(* IEC 61131-3 sources: 2026_Projet_YGO_ExcavatriceDragage/TOOLS/TEST_AUTO_CI/RESULTS/C_DIAG_RESEAUX/tests, 4 files *)

(* ---- test_fb_autoresettransientdiag.st ---- *)
(* =========================================================================
   FB_AutoResetTransientDiag — preuve isolee (T352, parent T278)
   =========================================================================
   Pourquoi ce fichier existe : T278 a livre le FB et son cablage SANS aucun
   test unitaire, et ses deux entrees d'autorisation StartupEnable /
   PowerRearmEnable ont ete cablees sur deux booleens d'une GVL de simulation
   valant FALSE par defaut et sans aucun ecrivain (PRG_02_Acquisition.st:225-226,
   GVL_Simulation.st:106-107). Consequence mesuree sur machine reelle : State
   reste bloque a 0, Phase ne passe jamais a 1 ni a 2, ResetPulse ne bouge
   jamais. Ces cas prouvent que la logique INTERNE du FB est saine des que les
   deux entrees valent TRUE — le defaut etait donc bien en amont du FB.

   Identifiants TC-T352-xxx : cas d'execution rattaches a la tache T352. Ils ne
   prennent AUCUN identifiant TC-P12 du catalogue AF-12 : ce catalogue s'arrete
   a TC-P12-050 et un TC-P12-060 a ete explicitement REFUSE par l'humain
   (AF_Partie-12_Fonction_Diagnostic_v1.4.md, ligne 348).

   Ce fichier prouve des comportements OBSERVABLES par les sorties publiques
   (ResetPulse, SequenceActive, Lockout, Cancelled, Phase, AttemptCount) :
   State et StartupStarted sont des VAR privees, non lisibles de l'exterieur.

   Gardes de securite couvertes, jamais affaiblies :
     FB_AutoResetTransientDiag.st:70  SafeCommon = EmergencyChainClosed AND
                                      NOT PowerCutOffActive AND NOT MotionActive
     FB_AutoResetTransientDiag.st:122 annulation immediate si SafeCommon tombe
   ========================================================================= *)

SETUP
VAR
    FB : FB_AutoResetTransientDiag;
END_VAR
END_SETUP

(* -------------------------------------------------------------------------
   Cas nominal : demarrage, stabilisation, impulsion unique, verrouillage.
   C'est exactement le scenario que l'observateur ne voyait jamais sur machine.
   ------------------------------------------------------------------------- *)
TEST 'TC-T352-001 Demarrage par defaut : Phase 1, impulsion apres stabilisation, verrouillage'
    (* Scan 0 : conditions nominales, contacteur au repos -> la sequence demarre *)
    FB(Enable := TRUE,
       StartupEnable := TRUE,
       PowerRearmEnable := TRUE,
       EmergencyChainClosed := TRUE,
       PowerContactorEngaged := FALSE,
       PowerCutOffActive := FALSE,
       MotionActive := FALSE,
       DiagnosticsStable := TRUE,
       Cfg_MaxAttempts := 1,
       Cfg_StabilizationTime := T#1s,
       Cfg_InterAttemptTime := T#1s);
    ASSERT_TRUE(FB.SequenceActive, 'StartupEnable=TRUE -> sequence active des le 1er scan');
    ASSERT_EQ(FB.Phase, 1, 'Phase 1 = sequence de demarrage engagee');

    (* Scan 1 : aucune impulsion, la stabilisation est en cours *)
    FB(Enable := TRUE, StartupEnable := TRUE, PowerRearmEnable := TRUE,
       EmergencyChainClosed := TRUE, PowerContactorEngaged := FALSE,
       PowerCutOffActive := FALSE, MotionActive := FALSE, DiagnosticsStable := TRUE,
       Cfg_MaxAttempts := 1, Cfg_StabilizationTime := T#1s, Cfg_InterAttemptTime := T#1s);
    ASSERT_FALSE(FB.ResetPulse, 'Aucune impulsion avant Cfg_StabilizationTime');

    (* Scan 2 : 1 s ecoulee -> impulsion unique puis verrouillage (MaxAttempts=1) *)
    ADVANCE_TIME(1000000000);
    FB(Enable := TRUE, StartupEnable := TRUE, PowerRearmEnable := TRUE,
       EmergencyChainClosed := TRUE, PowerContactorEngaged := FALSE,
       PowerCutOffActive := FALSE, MotionActive := FALSE, DiagnosticsStable := TRUE,
       Cfg_MaxAttempts := 1, Cfg_StabilizationTime := T#1s, Cfg_InterAttemptTime := T#1s);
    ASSERT_TRUE(FB.ResetPulse, 'Apres 1 s de stabilisation -> ResetPulse=TRUE');
    ASSERT_EQ(FB.AttemptCount, 1, 'Une seule impulsion emise');
    ASSERT_TRUE(FB.Lockout, 'MaxAttempts=1 atteint -> Lockout=TRUE');
    ASSERT_EQ(FB.Phase, 3, 'Phase 3 = salve terminee, attente d''un nouvel evenement');

    (* Scan 3 : impulsion d'un seul scan, puis retour au repos verrouille *)
    FB(Enable := TRUE, StartupEnable := TRUE, PowerRearmEnable := TRUE,
       EmergencyChainClosed := TRUE, PowerContactorEngaged := FALSE,
       PowerCutOffActive := FALSE, MotionActive := FALSE, DiagnosticsStable := TRUE,
       Cfg_MaxAttempts := 1, Cfg_StabilizationTime := T#1s, Cfg_InterAttemptTime := T#1s);
    ASSERT_FALSE(FB.ResetPulse, 'ResetPulse est impulsionnel : FALSE au scan suivant');
    ASSERT_TRUE(FB.Lockout, 'Lockout persiste apres la salve');
    ASSERT_FALSE(FB.SequenceActive, 'Sequence terminee');
END_TEST

(* -------------------------------------------------------------------------
   Le second chemin d'entree, inerte tant que PowerRearmEnable valait FALSE :
   phase 2 declenchee EXCLUSIVEMENT sur front du retour contacteur.
   ------------------------------------------------------------------------- *)
TEST 'TC-T352-002 Post-rearmement : Phase 2 sur front contacteur, impulsion puis verrouillage'
    (* Scan 0 : contacteur au repos, phase demarrage volontairement desactivee *)
    FB(Enable := TRUE,
       StartupEnable := FALSE,
       PowerRearmEnable := TRUE,
       EmergencyChainClosed := TRUE,
       PowerContactorEngaged := FALSE,
       PowerCutOffActive := FALSE,
       MotionActive := FALSE,
       DiagnosticsStable := TRUE,
       Cfg_MaxAttempts := 1,
       Cfg_StabilizationTime := T#1s,
       Cfg_InterAttemptTime := T#1s);
    ASSERT_FALSE(FB.SequenceActive, 'Aucun evenement -> sequence au repos');

    (* Scan 1 : front montant du contacteur -> phase post-rearmement *)
    FB(Enable := TRUE, StartupEnable := FALSE, PowerRearmEnable := TRUE,
       EmergencyChainClosed := TRUE, PowerContactorEngaged := TRUE,
       PowerCutOffActive := FALSE, MotionActive := FALSE, DiagnosticsStable := TRUE,
       Cfg_MaxAttempts := 1, Cfg_StabilizationTime := T#1s, Cfg_InterAttemptTime := T#1s);
    ASSERT_TRUE(FB.SequenceActive, 'Front contacteur -> sequence post-rearmement engagee');
    ASSERT_EQ(FB.Phase, 2, 'Phase 2 = sequence post-rearmement');
    ASSERT_FALSE(FB.ResetPulse, 'Impulsion differee apres stabilisation');

    (* Scan 2 : stabilisation ecoulee -> impulsion puis verrouillage *)
    ADVANCE_TIME(1000000000);
    FB(Enable := TRUE, StartupEnable := FALSE, PowerRearmEnable := TRUE,
       EmergencyChainClosed := TRUE, PowerContactorEngaged := TRUE,
       PowerCutOffActive := FALSE, MotionActive := FALSE, DiagnosticsStable := TRUE,
       Cfg_MaxAttempts := 1, Cfg_StabilizationTime := T#1s, Cfg_InterAttemptTime := T#1s);
    ASSERT_TRUE(FB.ResetPulse, 'Apres stabilisation post-rearmement -> ResetPulse=TRUE');
    ASSERT_EQ(FB.AttemptCount, 1, 'Une impulsion emise');
    ASSERT_TRUE(FB.Lockout, 'Salve epuisee -> Lockout=TRUE');
END_TEST

(* -------------------------------------------------------------------------
   Gardes de securite : aucune impulsion ne doit sortir. Les trois composantes
   de SafeCommon sont testees separement, chacune suffit a interdire la salve.
   ------------------------------------------------------------------------- *)
TEST 'TC-T352-003 Gardes safety : chaine AU ouverte, coupure puissance, mouvement actif'
    (* Chaine AU ouverte : EmergencyChainClosed=FALSE *)
    FB(Enable := TRUE, StartupEnable := TRUE, PowerRearmEnable := TRUE,
       EmergencyChainClosed := FALSE, PowerContactorEngaged := FALSE,
       PowerCutOffActive := FALSE, MotionActive := FALSE, DiagnosticsStable := TRUE,
       Cfg_MaxAttempts := 3, Cfg_StabilizationTime := T#1s, Cfg_InterAttemptTime := T#1s);
    ASSERT_FALSE(FB.SequenceActive, 'Chaine AU ouverte -> aucune sequence');
    ASSERT_FALSE(FB.ResetPulse, 'Chaine AU ouverte -> aucune impulsion');

    (* Coupure puissance active : PowerCutOffActive=TRUE *)
    FB(Enable := TRUE, StartupEnable := TRUE, PowerRearmEnable := TRUE,
       EmergencyChainClosed := TRUE, PowerContactorEngaged := FALSE,
       PowerCutOffActive := TRUE, MotionActive := FALSE, DiagnosticsStable := TRUE,
       Cfg_MaxAttempts := 3, Cfg_StabilizationTime := T#1s, Cfg_InterAttemptTime := T#1s);
    ASSERT_FALSE(FB.SequenceActive, 'Coupure puissance active -> aucune sequence');

    (* Mouvement actif : MotionActive=TRUE *)
    FB(Enable := TRUE, StartupEnable := TRUE, PowerRearmEnable := TRUE,
       EmergencyChainClosed := TRUE, PowerContactorEngaged := FALSE,
       PowerCutOffActive := FALSE, MotionActive := TRUE, DiagnosticsStable := TRUE,
       Cfg_MaxAttempts := 3, Cfg_StabilizationTime := T#1s, Cfg_InterAttemptTime := T#1s);
    ASSERT_FALSE(FB.SequenceActive, 'Mouvement actif -> aucune sequence');

    (* Le temps qui passe ne force rien : meme apres 5 s, toujours aucune impulsion *)
    ADVANCE_TIME(5000000000);
    FB(Enable := TRUE, StartupEnable := TRUE, PowerRearmEnable := TRUE,
       EmergencyChainClosed := TRUE, PowerContactorEngaged := FALSE,
       PowerCutOffActive := FALSE, MotionActive := TRUE, DiagnosticsStable := TRUE,
       Cfg_MaxAttempts := 3, Cfg_StabilizationTime := T#1s, Cfg_InterAttemptTime := T#1s);
    ASSERT_FALSE(FB.ResetPulse, 'Garde safety invalide -> ResetPulse reste FALSE malgre le temps');
    ASSERT_EQ(FB.AttemptCount, 0, 'Aucune tentative consommee sous garde invalide');

    (* Diagnostics reseau instables : la stabilisation ne progresse pas *)
    FB(Enable := TRUE, StartupEnable := TRUE, PowerRearmEnable := TRUE,
       EmergencyChainClosed := TRUE, PowerContactorEngaged := FALSE,
       PowerCutOffActive := FALSE, MotionActive := FALSE, DiagnosticsStable := FALSE,
       Cfg_MaxAttempts := 3, Cfg_StabilizationTime := T#1s, Cfg_InterAttemptTime := T#1s);
    ASSERT_EQ(FB.Phase, 1, 'Sequence engagee mais bloquee en phase 1');
    ADVANCE_TIME(5000000000);
    FB(Enable := TRUE, StartupEnable := TRUE, PowerRearmEnable := TRUE,
       EmergencyChainClosed := TRUE, PowerContactorEngaged := FALSE,
       PowerCutOffActive := FALSE, MotionActive := FALSE, DiagnosticsStable := FALSE,
       Cfg_MaxAttempts := 3, Cfg_StabilizationTime := T#1s, Cfg_InterAttemptTime := T#1s);
    ASSERT_FALSE(FB.ResetPulse, 'Diagnostics instables -> aucune impulsion');
    ASSERT_EQ(FB.AttemptCount, 0, 'Aucune tentative consommee sans diagnostics stables');
END_TEST

(* -------------------------------------------------------------------------
   Annulation en cours de sequence : la garde retombe pendant la salve.
   ------------------------------------------------------------------------- *)
TEST 'TC-T352-004 Annulation : chute de la garde pendant la sequence -> Cancelled + Lockout'
    FB(Enable := TRUE, StartupEnable := TRUE, PowerRearmEnable := TRUE,
       EmergencyChainClosed := TRUE, PowerContactorEngaged := FALSE,
       PowerCutOffActive := FALSE, MotionActive := FALSE, DiagnosticsStable := TRUE,
       Cfg_MaxAttempts := 3, Cfg_StabilizationTime := T#1s, Cfg_InterAttemptTime := T#1s);
    ASSERT_EQ(FB.Phase, 1, 'Sequence engagee');

    (* L'AU s'ouvre pendant la salve -> annulation immediate *)
    ADVANCE_TIME(500000000);
    FB(Enable := TRUE, StartupEnable := TRUE, PowerRearmEnable := TRUE,
       EmergencyChainClosed := FALSE, PowerContactorEngaged := FALSE,
       PowerCutOffActive := FALSE, MotionActive := FALSE, DiagnosticsStable := TRUE,
       Cfg_MaxAttempts := 3, Cfg_StabilizationTime := T#1s, Cfg_InterAttemptTime := T#1s);
    ASSERT_TRUE(FB.Cancelled, 'Garde tombee en cours de sequence -> Cancelled=TRUE');
    ASSERT_TRUE(FB.Lockout, 'Salve annulee -> Lockout=TRUE');
    ASSERT_FALSE(FB.ResetPulse, 'Annulation -> aucune impulsion');
    ASSERT_FALSE(FB.SequenceActive, 'Sequence interrompue');
    ASSERT_EQ(FB.Phase, 3, 'Phase 3 = verrouillage apres annulation');
END_TEST

(* -------------------------------------------------------------------------
   Borne haute : 3 impulsions espacees de Cfg_InterAttemptTime, puis lockout.
   Cadence reelle du FB : impulsion (etat 3) -> scan d'intervalle (retour etat 1)
   -> redemarrage de la stabilisation -> impulsion suivante.
   ------------------------------------------------------------------------- *)
TEST 'TC-T352-005 Borne haute : 3 impulsions espacees puis verrouillage definitif'
    FB(Enable := TRUE, StartupEnable := TRUE, PowerRearmEnable := TRUE,
       EmergencyChainClosed := TRUE, PowerContactorEngaged := FALSE,
       PowerCutOffActive := FALSE, MotionActive := FALSE, DiagnosticsStable := TRUE,
       Cfg_MaxAttempts := 3, Cfg_StabilizationTime := T#1s, Cfg_InterAttemptTime := T#1s);
    ASSERT_EQ(FB.Phase, 1, 'Sequence engagee');

    (* Impulsion 1 *)
    ADVANCE_TIME(1000000000);
    FB(Enable := TRUE, StartupEnable := TRUE, PowerRearmEnable := TRUE,
       EmergencyChainClosed := TRUE, PowerContactorEngaged := FALSE,
       PowerCutOffActive := FALSE, MotionActive := FALSE, DiagnosticsStable := TRUE,
       Cfg_MaxAttempts := 3, Cfg_StabilizationTime := T#1s, Cfg_InterAttemptTime := T#1s);
    ASSERT_TRUE(FB.ResetPulse, 'Impulsion 1 sur 3');
    ASSERT_EQ(FB.AttemptCount, 1, 'Compteur a 1');
    ASSERT_FALSE(FB.Lockout, 'Salve non epuisee -> aucun verrouillage');

    (* Intervalle : la tempo inter-impulsions ramene la sequence en phase 1 *)
    ADVANCE_TIME(1000000000);
    FB(Enable := TRUE, StartupEnable := TRUE, PowerRearmEnable := TRUE,
       EmergencyChainClosed := TRUE, PowerContactorEngaged := FALSE,
       PowerCutOffActive := FALSE, MotionActive := FALSE, DiagnosticsStable := TRUE,
       Cfg_MaxAttempts := 3, Cfg_StabilizationTime := T#1s, Cfg_InterAttemptTime := T#1s);
    ASSERT_FALSE(FB.ResetPulse, 'Intervalle inter-impulsions respecte');
    ASSERT_EQ(FB.AttemptCount, 1, 'Compteur inchange pendant l''intervalle');
    ASSERT_EQ(FB.Phase, 1, 'Retour en phase 1 pour la tentative suivante');

    (* Redemarrage de la stabilisation puis impulsion 2 *)
    ADVANCE_TIME(1000000000);
    FB(Enable := TRUE, StartupEnable := TRUE, PowerRearmEnable := TRUE,
       EmergencyChainClosed := TRUE, PowerContactorEngaged := FALSE,
       PowerCutOffActive := FALSE, MotionActive := FALSE, DiagnosticsStable := TRUE,
       Cfg_MaxAttempts := 3, Cfg_StabilizationTime := T#1s, Cfg_InterAttemptTime := T#1s);
    ASSERT_FALSE(FB.ResetPulse, 'Stabilisation redemarree : pas d''impulsion immediate');

    ADVANCE_TIME(1000000000);
    FB(Enable := TRUE, StartupEnable := TRUE, PowerRearmEnable := TRUE,
       EmergencyChainClosed := TRUE, PowerContactorEngaged := FALSE,
       PowerCutOffActive := FALSE, MotionActive := FALSE, DiagnosticsStable := TRUE,
       Cfg_MaxAttempts := 3, Cfg_StabilizationTime := T#1s, Cfg_InterAttemptTime := T#1s);
    ASSERT_TRUE(FB.ResetPulse, 'Impulsion 2 sur 3');
    ASSERT_EQ(FB.AttemptCount, 2, 'Compteur a 2');
    ASSERT_FALSE(FB.Lockout, 'Salve non epuisee -> aucun verrouillage');

    (* Intervalle puis impulsion 3, qui sature la borne *)
    ADVANCE_TIME(1000000000);
    FB(Enable := TRUE, StartupEnable := TRUE, PowerRearmEnable := TRUE,
       EmergencyChainClosed := TRUE, PowerContactorEngaged := FALSE,
       PowerCutOffActive := FALSE, MotionActive := FALSE, DiagnosticsStable := TRUE,
       Cfg_MaxAttempts := 3, Cfg_StabilizationTime := T#1s, Cfg_InterAttemptTime := T#1s);
    ASSERT_FALSE(FB.ResetPulse, 'Intervalle inter-impulsions respecte (2)');

    ADVANCE_TIME(1000000000);
    FB(Enable := TRUE, StartupEnable := TRUE, PowerRearmEnable := TRUE,
       EmergencyChainClosed := TRUE, PowerContactorEngaged := FALSE,
       PowerCutOffActive := FALSE, MotionActive := FALSE, DiagnosticsStable := TRUE,
       Cfg_MaxAttempts := 3, Cfg_StabilizationTime := T#1s, Cfg_InterAttemptTime := T#1s);
    ASSERT_FALSE(FB.ResetPulse, 'Stabilisation redemarree : pas d''impulsion immediate (2)');

    ADVANCE_TIME(1000000000);
    FB(Enable := TRUE, StartupEnable := TRUE, PowerRearmEnable := TRUE,
       EmergencyChainClosed := TRUE, PowerContactorEngaged := FALSE,
       PowerCutOffActive := FALSE, MotionActive := FALSE, DiagnosticsStable := TRUE,
       Cfg_MaxAttempts := 3, Cfg_StabilizationTime := T#1s, Cfg_InterAttemptTime := T#1s);
    ASSERT_TRUE(FB.ResetPulse, 'Impulsion 3 sur 3');
    ASSERT_EQ(FB.AttemptCount, 3, 'Compteur a 3');
    ASSERT_TRUE(FB.Lockout, 'Borne haute atteinte -> verrouillage');
    ASSERT_EQ(FB.Phase, 3, 'Phase 3 apres salve complete');

    (* Le temps ne relance rien : seul un nouvel evenement rearme la salve *)
    ADVANCE_TIME(10000000000);
    FB(Enable := TRUE, StartupEnable := TRUE, PowerRearmEnable := TRUE,
       EmergencyChainClosed := TRUE, PowerContactorEngaged := FALSE,
       PowerCutOffActive := FALSE, MotionActive := FALSE, DiagnosticsStable := TRUE,
       Cfg_MaxAttempts := 3, Cfg_StabilizationTime := T#1s, Cfg_InterAttemptTime := T#1s);
    ASSERT_FALSE(FB.ResetPulse, 'Aucune 4e impulsion');
    ASSERT_EQ(FB.AttemptCount, 3, 'Compteur fige a la borne');
    ASSERT_TRUE(FB.Lockout, 'Verrouillage conserve');
END_TEST

(* -------------------------------------------------------------------------
   Neutralisation : Enable=FALSE remet le service au repos.
   ------------------------------------------------------------------------- *)
TEST 'TC-T352-006 Neutralisation : Enable=FALSE -> service remis au repos'
    FB(Enable := TRUE, StartupEnable := TRUE, PowerRearmEnable := TRUE,
       EmergencyChainClosed := TRUE, PowerContactorEngaged := FALSE,
       PowerCutOffActive := FALSE, MotionActive := FALSE, DiagnosticsStable := TRUE,
       Cfg_MaxAttempts := 3, Cfg_StabilizationTime := T#1s, Cfg_InterAttemptTime := T#1s);
    ASSERT_TRUE(FB.SequenceActive, 'Sequence engagee avant neutralisation');

    FB(Enable := FALSE, StartupEnable := TRUE, PowerRearmEnable := TRUE,
       EmergencyChainClosed := TRUE, PowerContactorEngaged := FALSE,
       PowerCutOffActive := FALSE, MotionActive := FALSE, DiagnosticsStable := TRUE,
       Cfg_MaxAttempts := 3, Cfg_StabilizationTime := T#1s, Cfg_InterAttemptTime := T#1s);
    ASSERT_FALSE(FB.SequenceActive, 'Enable=FALSE -> sequence neutralisee');
    ASSERT_FALSE(FB.Lockout, 'Enable=FALSE -> verrouillage efface');
    ASSERT_EQ(FB.Phase, 0, 'Enable=FALSE -> retour au repos');
    ASSERT_EQ(FB.AttemptCount, 0, 'Enable=FALSE -> compteur remis a zero');
    ASSERT_FALSE(FB.ResetPulse, 'Enable=FALSE -> aucune impulsion');
END_TEST

(* ---- test_fb_diag_canopen.st ---- *)
SETUP
VAR
    FB : FB_Diag_CanOpen;
END_VAR
END_SETUP

TEST 'TC-P03-001 Dynamique Enable : neutralisation initiale, transition Ready au repos, puis coupure'
    (* Scan 0 : Enable=FALSE -> Diagnostic desactive *)
    FB(Enable := FALSE, CANbusStateRaw := 2, DeviceJoystickStateRaw := DEVICE_STATE.RUNNING);
    ASSERT_FALSE(FB.Ready, 'Enable=FALSE -> Ready=FALSE (neutralise)');
    ASSERT_EQ(FB.DeviceCanOpenMaster.State, E_Diag_State.DISABLED, 'State doit etre DISABLED sans Enable');

    ADVANCE_TIME(10000000);

    (* Scan 1 : Enable=TRUE -> Diagnostic pret et actif *)
    FB(Enable := TRUE, CANbusStateRaw := 2, DeviceJoystickStateRaw := DEVICE_STATE.RUNNING,
       SimBypassActive := FALSE, NetworkBypassActive := FALSE);
    ASSERT_TRUE(FB.Ready, 'Enable=TRUE -> Ready=TRUE (nominal)');
    ASSERT_EQ(FB.DeviceCanOpenMaster.State, E_Diag_State.READY, 'State doit etre READY');

    ADVANCE_TIME(10000000);

    (* Scan 2 : Enable=FALSE -> Re-neutralisation *)
    FB(Enable := FALSE, CANbusStateRaw := 2, DeviceJoystickStateRaw := DEVICE_STATE.RUNNING);
    ASSERT_FALSE(FB.Ready, 'Enable=FALSE -> Ready retombe a FALSE');
    ASSERT_EQ(FB.DeviceCanOpenMaster.State, E_Diag_State.DISABLED, 'State retombe a DISABLED');
END_TEST

TEST 'TC-P12-001 CanOpen : surveillance bus et esclave'
    FB(Enable := TRUE, CANbusStateRaw := 2, DeviceJoystickStateRaw := DEVICE_STATE.RUNNING,
       SimBypassActive := FALSE, NetworkBypassActive := FALSE);
    ASSERT_TRUE(FB.Ready, 'Bus et esclave sains');
    ASSERT_FALSE(FB.DeviceCanOpenMaster.Error, 'Aucune erreur bus maitre');
    ASSERT_FALSE(FB.DeviceJoystick.Error, 'Aucune erreur joystick');
END_TEST

(* =========================================================================
   AF-12 — Diagnostic : TC-P12-040 (bypass sim/reseau vs etat reel)
   ========================================================================= *)

TEST 'TC-P12-040 CanOpen : bypass sim/reseau vs etat reel (READY/SIMULATED/DISABLED)'
    (* Reel RUNNING sans bypass -> READY *)
    FB(Enable := TRUE, CANbusStateRaw := 2, DeviceJoystickStateRaw := DEVICE_STATE.RUNNING,
       SimBypassActive := FALSE, NetworkBypassActive := FALSE);
    ASSERT_EQ(FB.DeviceJoystick.State, E_Diag_State.READY, 'Reel RUNNING sans bypass -> READY');

    (* Bypass sans device reel -> SIMULATED *)
    FB(Enable := TRUE, CANbusStateRaw := 0, DeviceJoystickStateRaw := DEVICE_STATE.STOPPED,
       SimBypassActive := TRUE, NetworkBypassActive := FALSE);
    ASSERT_EQ(FB.DeviceJoystick.State, E_Diag_State.SIMULATED, 'Bypass sans device reel -> SIMULATED');

    (* Ni l un ni l autre -> ERROR (fiche attend INIT, code produit ERROR -- ecart documente AF12 TBD) *)
    FB(Enable := TRUE, CANbusStateRaw := 0, DeviceJoystickStateRaw := DEVICE_STATE.STOPPED,
       SimBypassActive := FALSE, NetworkBypassActive := FALSE);
    ASSERT_EQ(FB.DeviceJoystick.State, E_Diag_State.ERROR, 'Ni bypass ni reel -> ERROR (ecart fiche INIT)');

    (* Enable=FALSE prioritaire -> DISABLED *)
    FB(Enable := FALSE, CANbusStateRaw := 2, DeviceJoystickStateRaw := DEVICE_STATE.RUNNING);
    ASSERT_EQ(FB.DeviceJoystick.State, E_Diag_State.DISABLED, 'Enable=FALSE -> DISABLED');
END_TEST

(* ---- test_fb_diag_ethercat.st ---- *)
SETUP
VAR
    FB : FB_Diag_Ethercat;
    (* Temoin de l'invariance T359 : meme sequence, SANS jamais activer ResetTransient.
       Toute difference entre FB et FBCtrl signerait un effet reel du pulse d'auto-acquittement. *)
    FBCtrl : FB_Diag_Ethercat;
END_VAR
END_SETUP

TEST 'TC-P03-001 Dynamique Enable : neutralisation initiale, transition Ready au repos, puis coupure'
    (* Scan 0 : Enable=FALSE -> Diagnostic desactive *)
    FB(Enable := FALSE, DeviceVariateurStateRaw := DEVICE_STATE.RUNNING,
       DeviceEncoderM1StateRaw := DEVICE_STATE.RUNNING, DeviceEncoderM2StateRaw := DEVICE_STATE.RUNNING);
    ASSERT_FALSE(FB.Ready, 'Enable=FALSE -> Ready=FALSE');
    ASSERT_EQ(FB.DeviceEthercatMaster.State, E_Diag_State.DISABLED, 'State=DISABLED');

    ADVANCE_TIME(10000000);

    (* Scan 1 : Enable=TRUE -> Diagnostic actif *)
    FB(Enable := TRUE, DeviceVariateurStateRaw := DEVICE_STATE.RUNNING,
       DeviceEncoderM1StateRaw := DEVICE_STATE.RUNNING, DeviceEncoderM2StateRaw := DEVICE_STATE.RUNNING,
       NetworkBypassActive := FALSE);
    ASSERT_TRUE(FB.Ready, 'Enable=TRUE -> Ready=TRUE');
    ASSERT_EQ(FB.DeviceEthercatMaster.State, E_Diag_State.READY, 'State=READY');

    ADVANCE_TIME(10000000);

    (* Scan 2 : Enable=FALSE -> Re-neutralisation *)
    FB(Enable := FALSE, DeviceVariateurStateRaw := DEVICE_STATE.RUNNING,
       DeviceEncoderM1StateRaw := DEVICE_STATE.RUNNING, DeviceEncoderM2StateRaw := DEVICE_STATE.RUNNING);
    ASSERT_FALSE(FB.Ready, 'Coupure -> Ready retombe a FALSE');
    ASSERT_EQ(FB.DeviceEthercatMaster.State, E_Diag_State.DISABLED, 'State retombe a DISABLED');
END_TEST

TEST 'TC-P12-010 EtherCAT : surveillance maitre et esclaves'
    FB(Enable := TRUE, DeviceVariateurStateRaw := DEVICE_STATE.RUNNING,
       DeviceEncoderM1StateRaw := DEVICE_STATE.RUNNING, DeviceEncoderM2StateRaw := DEVICE_STATE.RUNNING,
       NetworkBypassActive := FALSE);
    ASSERT_TRUE(FB.Ready, 'EtherCAT pret');
    ASSERT_FALSE(FB.DeviceEthercatMaster.Error, 'Pas d erreur bus');
    ASSERT_FALSE(FB.DeviceEncoderM1.Error, 'Pas d erreur encoder M1');
END_TEST

(* =========================================================================
   AF-12 — Diagnostic : TC-P12-030 (synthèse par device) & TC-P12-040 (bypass)
   ========================================================================= *)

TEST 'TC-P12-030 EtherCAT : State != RUNNING par device -> bits ErrorId + Error global'
    (* Variateur M3 hors RUNNING -> bit 4 (16#0010), M1/M2 sains *)
    FB(Enable := TRUE, DeviceVariateurStateRaw := DEVICE_STATE.STOPPED,
       DeviceEncoderM1StateRaw := DEVICE_STATE.RUNNING, DeviceEncoderM2StateRaw := DEVICE_STATE.RUNNING,
       NetworkBypassActive := FALSE);
    ASSERT_TRUE(FB.DeviceVariateur.Error, 'Variateur hors RUNNING -> Error=TRUE');
    ASSERT_EQ(FB.DeviceVariateur.ErrorId, 16#0010, 'Variateur -> ErrorId bit 4 (16#0010)');
    ASSERT_FALSE(FB.DeviceEncoderM1.Error, 'M1 sain -> pas d erreur');
    ASSERT_FALSE(FB.DeviceEncoderM2.Error, 'M2 sain -> pas d erreur');
    ASSERT_TRUE(FB.DeviceEthercatMaster.Error, 'Un device en defaut -> Error maitre=TRUE');

    (* M1 hors RUNNING -> bit 5 (16#0020), variateur/M2 sains *)
    FB(Enable := TRUE, DeviceVariateurStateRaw := DEVICE_STATE.RUNNING,
       DeviceEncoderM1StateRaw := DEVICE_STATE.STOPPED, DeviceEncoderM2StateRaw := DEVICE_STATE.RUNNING,
       NetworkBypassActive := FALSE);
    ASSERT_TRUE(FB.DeviceEncoderM1.Error, 'M1 hors RUNNING -> Error=TRUE');
    ASSERT_EQ(FB.DeviceEncoderM1.ErrorId, 16#0020, 'M1 -> ErrorId bit 5 (16#0020)');
    ASSERT_FALSE(FB.DeviceVariateur.Error, 'Variateur sain -> pas d erreur');

    (* M2 hors RUNNING -> 16#0030 (bug T159 documente, pas 16#0040) *)
    FB(Enable := TRUE, DeviceVariateurStateRaw := DEVICE_STATE.RUNNING,
       DeviceEncoderM1StateRaw := DEVICE_STATE.RUNNING, DeviceEncoderM2StateRaw := DEVICE_STATE.STOPPED,
       NetworkBypassActive := FALSE);
    ASSERT_TRUE(FB.DeviceEncoderM2.Error, 'M2 hors RUNNING -> Error=TRUE');
    ASSERT_EQ(FB.DeviceEncoderM2.ErrorId, 16#0030, 'M2 -> ErrorId 16#0030 (bug T159 documente)');
END_TEST

TEST 'TC-P12-040 EtherCAT : bypass sim/reseau vs etat reel (READY/SIMULATED/DISABLED)'
    (* Reel RUNNING sans bypass -> READY *)
    FB(Enable := TRUE, DeviceVariateurStateRaw := DEVICE_STATE.RUNNING,
       DeviceEncoderM1StateRaw := DEVICE_STATE.RUNNING, DeviceEncoderM2StateRaw := DEVICE_STATE.RUNNING,
       NetworkBypassActive := FALSE);
    ASSERT_EQ(FB.DeviceVariateur.State, E_Diag_State.READY, 'Reel RUNNING sans bypass -> READY');

    (* Bypass sans device reel -> SIMULATED *)
    FB(Enable := TRUE, DeviceVariateurStateRaw := DEVICE_STATE.STOPPED,
       DeviceEncoderM1StateRaw := DEVICE_STATE.RUNNING, DeviceEncoderM2StateRaw := DEVICE_STATE.RUNNING,
       NetworkBypassActive := TRUE);
    ASSERT_EQ(FB.DeviceVariateur.State, E_Diag_State.SIMULATED, 'Bypass sans device reel -> SIMULATED');

    (* Ni l un ni l autre -> ERROR (fiche attend INIT, code produit ERROR -- ecart documente AF12 TBD) *)
    FB(Enable := TRUE, DeviceVariateurStateRaw := DEVICE_STATE.STOPPED,
       DeviceEncoderM1StateRaw := DEVICE_STATE.RUNNING, DeviceEncoderM2StateRaw := DEVICE_STATE.RUNNING,
       NetworkBypassActive := FALSE);
    ASSERT_EQ(FB.DeviceVariateur.State, E_Diag_State.ERROR, 'Ni bypass ni reel -> ERROR (ecart fiche INIT)');

    (* Enable=FALSE prioritaire -> DISABLED *)
    FB(Enable := FALSE, DeviceVariateurStateRaw := DEVICE_STATE.RUNNING,
       DeviceEncoderM1StateRaw := DEVICE_STATE.RUNNING, DeviceEncoderM2StateRaw := DEVICE_STATE.RUNNING);
    ASSERT_EQ(FB.DeviceVariateur.State, E_Diag_State.DISABLED, 'Enable=FALSE -> DISABLED');
END_TEST

(* =========================================================================
   T359 — PREUVE QUE L'AUTO-ACQUITTEMENT ResetTransient EST UN NO-OP
   =========================================================================
   OBJET DE LA PREUVE (aucun correctif ici, preuve AVANT correctif) : le service
   d'auto-acquittement borne (FB_AutoResetTransientDiag) produit bien une impulsion
   ResetTransient, mais cette impulsion n'a AUCUN effet observable sur les bits de
   diagnostic. Demonstration par trois faits :

   1. ORDRE DE SCAN (FB_Diag_Ethercat.st) : le bloc reset (lignes 103-119, dont
      ResetTransient en 106-112) s'execute AVANT le bloc « Diagnostic par equipement »
      (lignes 123-152) qui contient l'effacement automatique `AND 16#FFEF` (ligne 131),
      `16#FFDF` (141), `16#FFCF` (151). L'effet du pulse est donc ECRASE DANS LE MEME SCAN.

   2. L'effacement automatique est PREEXISTANT a T278 : le commit cb5ae5ea n'ajoute QUE
      la voie ResetTransient (git show cb5ae5ea -- CODE/C_DIAG_RESEAUX/FB_Diag_Ethercat.st
      ne contient ni 131, ni 141, ni 151). La fonctionnalite etait inoperante a sa
      conception, independamment des flags d'activation corriges en T352.

   3. INVARIANCE : ErrorId de fin de scan = f(OnlineEff) SEUL.
      - OnlineEff = TRUE  -> l'effacement automatique passe, que le pulse ait agi ou non ;
      - OnlineEff = FALSE -> la garde du pulse (`IF VariateurOnlineEff`) est fausse, le bit
        est pose a nouveau juste apres par la ligne 129.
      => ResetTransient ne peut rien changer. C'est ce que mesurent ces 3 tests, en
      comparant FB (avec pulse) et FBCtrl (sans pulse) EGAL A EGAL.
   ========================================================================= *)

TEST 'TC-T359-001 Invariance : une perte de liaison puis retour, pulse actif vs temoin sans pulse'
    (* Scan 0 : tout est en ligne, aucune impulsion *)
    FB(Enable := TRUE, DeviceVariateurStateRaw := DEVICE_STATE.RUNNING,
       DeviceEncoderM1StateRaw := DEVICE_STATE.RUNNING, DeviceEncoderM2StateRaw := DEVICE_STATE.RUNNING,
       NetworkBypassActive := FALSE, EcatBusBypassActive := FALSE, ResetTransient := FALSE);
    FBCtrl(Enable := TRUE, DeviceVariateurStateRaw := DEVICE_STATE.RUNNING,
       DeviceEncoderM1StateRaw := DEVICE_STATE.RUNNING, DeviceEncoderM2StateRaw := DEVICE_STATE.RUNNING,
       NetworkBypassActive := FALSE, EcatBusBypassActive := FALSE, ResetTransient := FALSE);
    ASSERT_EQ(FB.DeviceVariateur.ErrorId, 16#0000, 'Etat initial sain : ErrorId variateur nul');

    (* Scan 1 : PERTE DE LIAISON variateur -> le bit est pose *)
    FB(Enable := TRUE, DeviceVariateurStateRaw := DEVICE_STATE.STOPPED,
       DeviceEncoderM1StateRaw := DEVICE_STATE.RUNNING, DeviceEncoderM2StateRaw := DEVICE_STATE.RUNNING,
       NetworkBypassActive := FALSE, EcatBusBypassActive := FALSE, ResetTransient := FALSE);
    FBCtrl(Enable := TRUE, DeviceVariateurStateRaw := DEVICE_STATE.STOPPED,
       DeviceEncoderM1StateRaw := DEVICE_STATE.RUNNING, DeviceEncoderM2StateRaw := DEVICE_STATE.RUNNING,
       NetworkBypassActive := FALSE, EcatBusBypassActive := FALSE, ResetTransient := FALSE);
    ASSERT_EQ(FB.DeviceVariateur.ErrorId, 16#0010, 'Perte liaison variateur -> bit 16#0010 pose');
    ASSERT_FALSE(FB.DeviceVariateur.Online, 'Variateur hors ligne pendant la perte');

    (* Scan 2 : RETOUR DE LIAISON, front ResetTransient sur FB seul (FBCtrl reste sans pulse) *)
    FB(Enable := TRUE, DeviceVariateurStateRaw := DEVICE_STATE.RUNNING,
       DeviceEncoderM1StateRaw := DEVICE_STATE.RUNNING, DeviceEncoderM2StateRaw := DEVICE_STATE.RUNNING,
       NetworkBypassActive := FALSE, EcatBusBypassActive := FALSE, ResetTransient := TRUE);
    FBCtrl(Enable := TRUE, DeviceVariateurStateRaw := DEVICE_STATE.RUNNING,
       DeviceEncoderM1StateRaw := DEVICE_STATE.RUNNING, DeviceEncoderM2StateRaw := DEVICE_STATE.RUNNING,
       NetworkBypassActive := FALSE, EcatBusBypassActive := FALSE, ResetTransient := FALSE);

    (* Aucun scan n'expose « en ligne ET bit pose » : l'effacement automatique a deja agi *)
    ASSERT_TRUE(FB.DeviceVariateur.Online, 'Variateur de nouveau en ligne');
    ASSERT_EQ(FB.DeviceVariateur.ErrorId, 16#0000, 'Bit deja efface SANS le pulse (effacement auto ligne 131)');

    (* PREUVE D'INVARIANCE : le pulse ne change RIEN *)
    ASSERT_EQ(FB.DeviceVariateur.ErrorId, FBCtrl.DeviceVariateur.ErrorId,
              'INVARIANCE : ErrorId identique avec et sans ResetTransient');
    ASSERT_EQ(FB.DeviceVariateur.Error, FBCtrl.DeviceVariateur.Error,
              'INVARIANCE : Error identique avec et sans ResetTransient');
    ASSERT_EQ(FB.DeviceEthercatMaster.ErrorId, FBCtrl.DeviceEthercatMaster.ErrorId,
              'INVARIANCE : aucun effet sur le diagnostic maitre non plus');
END_TEST

TEST 'TC-T359-002 Invariance au timing de production : pulse 1 s APRES le retour de liaison'
    (* Scan 0 : tout en ligne *)
    FB(Enable := TRUE, DeviceVariateurStateRaw := DEVICE_STATE.RUNNING,
       DeviceEncoderM1StateRaw := DEVICE_STATE.RUNNING, DeviceEncoderM2StateRaw := DEVICE_STATE.RUNNING,
       NetworkBypassActive := FALSE, EcatBusBypassActive := FALSE, ResetTransient := FALSE);
    FBCtrl(Enable := TRUE, DeviceVariateurStateRaw := DEVICE_STATE.RUNNING,
       DeviceEncoderM1StateRaw := DEVICE_STATE.RUNNING, DeviceEncoderM2StateRaw := DEVICE_STATE.RUNNING,
       NetworkBypassActive := FALSE, EcatBusBypassActive := FALSE, ResetTransient := FALSE);

    (* Scan 1 : perte des DEUX codeurs *)
    FB(Enable := TRUE, DeviceVariateurStateRaw := DEVICE_STATE.RUNNING,
       DeviceEncoderM1StateRaw := DEVICE_STATE.STOPPED, DeviceEncoderM2StateRaw := DEVICE_STATE.STOPPED,
       NetworkBypassActive := FALSE, EcatBusBypassActive := FALSE, ResetTransient := FALSE);
    FBCtrl(Enable := TRUE, DeviceVariateurStateRaw := DEVICE_STATE.RUNNING,
       DeviceEncoderM1StateRaw := DEVICE_STATE.STOPPED, DeviceEncoderM2StateRaw := DEVICE_STATE.STOPPED,
       NetworkBypassActive := FALSE, EcatBusBypassActive := FALSE, ResetTransient := FALSE);
    ASSERT_EQ(FB.DeviceEncoderM1.ErrorId, 16#0020, 'Perte liaison codeur M1 -> bit 16#0020');
    ASSERT_EQ(FB.DeviceEncoderM2.ErrorId, 16#0030, 'Perte liaison codeur M2 -> bit 16#0030');

    (* Scan 2 : retour de liaison, PAS encore de pulse (comme sur machine : la sequence attend
       Cfg_StabilizationTime = 1 s avant d'emetre son impulsion) *)
    FB(Enable := TRUE, DeviceVariateurStateRaw := DEVICE_STATE.RUNNING,
       DeviceEncoderM1StateRaw := DEVICE_STATE.RUNNING, DeviceEncoderM2StateRaw := DEVICE_STATE.RUNNING,
       NetworkBypassActive := FALSE, EcatBusBypassActive := FALSE, ResetTransient := FALSE);
    FBCtrl(Enable := TRUE, DeviceVariateurStateRaw := DEVICE_STATE.RUNNING,
       DeviceEncoderM1StateRaw := DEVICE_STATE.RUNNING, DeviceEncoderM2StateRaw := DEVICE_STATE.RUNNING,
       NetworkBypassActive := FALSE, EcatBusBypassActive := FALSE, ResetTransient := FALSE);
    ASSERT_EQ(FB.DeviceEncoderM1.ErrorId, 16#0000, 'Codeur M1 deja efface au retour de liaison');
    ASSERT_EQ(FB.DeviceEncoderM2.ErrorId, 16#0000, 'Codeur M2 deja efface au retour de liaison');

    (* Scan 3 : 1 s plus tard, l'impulsion d'auto-acquittement arrive enfin *)
    ADVANCE_TIME(1000000000);
    FB(Enable := TRUE, DeviceVariateurStateRaw := DEVICE_STATE.RUNNING,
       DeviceEncoderM1StateRaw := DEVICE_STATE.RUNNING, DeviceEncoderM2StateRaw := DEVICE_STATE.RUNNING,
       NetworkBypassActive := FALSE, EcatBusBypassActive := FALSE, ResetTransient := TRUE);
    FBCtrl(Enable := TRUE, DeviceVariateurStateRaw := DEVICE_STATE.RUNNING,
       DeviceEncoderM1StateRaw := DEVICE_STATE.RUNNING, DeviceEncoderM2StateRaw := DEVICE_STATE.RUNNING,
       NetworkBypassActive := FALSE, EcatBusBypassActive := FALSE, ResetTransient := FALSE);
    ASSERT_EQ(FB.DeviceEncoderM1.ErrorId, FBCtrl.DeviceEncoderM1.ErrorId,
              'INVARIANCE : pulse tardif sans effet sur codeur M1');
    ASSERT_EQ(FB.DeviceEncoderM2.ErrorId, FBCtrl.DeviceEncoderM2.ErrorId,
              'INVARIANCE : pulse tardif sans effet sur codeur M2');
    ASSERT_EQ(FB.DeviceEthercatMaster.ErrorId, FBCtrl.DeviceEthercatMaster.ErrorId,
              'INVARIANCE : pulse tardif sans effet sur le maitre');
END_TEST

TEST 'TC-T359-003 La voie alternative « front Online » ne peut pas davantage agir sur le bit'
    (* Cette sequence prouve que le bit de liaison n'est JAMAIS observable a TRUE alors que
       l'equipement est en ligne : il n'existe donc aucun instant ou un pulse, meme declenche
       au scan exact du front Online, aurait quelque chose a effacer. *)
    FB(Enable := TRUE, DeviceVariateurStateRaw := DEVICE_STATE.STOPPED,
       DeviceEncoderM1StateRaw := DEVICE_STATE.STOPPED, DeviceEncoderM2StateRaw := DEVICE_STATE.STOPPED,
       NetworkBypassActive := FALSE, EcatBusBypassActive := FALSE, ResetTransient := FALSE);
    ASSERT_FALSE(FB.DeviceVariateur.Online, 'Hors ligne : bit pose, aucun pulse possible (garde OnlineEff)');
    ASSERT_EQ(FB.DeviceVariateur.ErrorId, 16#0010, 'Hors ligne : bit pose');

    (* Le scan EXACT du retour : Online passe a TRUE et le bit tombe dans le meme scan *)
    FB(Enable := TRUE, DeviceVariateurStateRaw := DEVICE_STATE.RUNNING,
       DeviceEncoderM1StateRaw := DEVICE_STATE.RUNNING, DeviceEncoderM2StateRaw := DEVICE_STATE.RUNNING,
       NetworkBypassActive := FALSE, EcatBusBypassActive := FALSE, ResetTransient := FALSE);
    ASSERT_TRUE(FB.DeviceVariateur.Online, 'Scan du front Online : variateur en ligne');
    ASSERT_EQ(FB.DeviceVariateur.ErrorId, 16#0000,
              'Scan du front Online : le bit est deja a 0 dans LE MEME scan — rien a effacer');

    (* Contre-epreuve du temoin : le pulse ACTIF sur ce meme scan ne peut pas faire mieux *)
    ADVANCE_TIME(10000000);
    FBCtrl(Enable := TRUE, DeviceVariateurStateRaw := DEVICE_STATE.RUNNING,
       DeviceEncoderM1StateRaw := DEVICE_STATE.RUNNING, DeviceEncoderM2StateRaw := DEVICE_STATE.RUNNING,
       NetworkBypassActive := FALSE, EcatBusBypassActive := FALSE, ResetTransient := TRUE);
    ASSERT_EQ(FBCtrl.DeviceVariateur.ErrorId, 16#0000,
              'Contre-epreuve : pulse au scan du front Online -> toujours 0, aucune valeur ajoutee');
END_TEST

(* ---- test_fb_diag_ihmheartbeat.st ---- *)
SETUP
VAR
    FB : FB_Diag_IhmHeartbeat;
END_VAR
END_SETUP

TEST 'TC-P03-001 Dynamique Enable : neutralisation initiale, transition HeartbeatIhmOk, puis coupure'
    (* Scan 0 : Enable=FALSE -> Diagnostic desactive *)
    FB(Enable := FALSE, TglHeartbeatIhm := FALSE, IhmTimeout := T#2s);
    ASSERT_FALSE(FB.HeartbeatIhmOk, 'Enable=FALSE -> HeartbeatIhmOk=FALSE');
    ASSERT_TRUE(FB.HeartbeatIhmTimeout, 'Enable=FALSE -> HeartbeatIhmTimeout=TRUE');

    ADVANCE_TIME(10000000);

    (* Scan 1 : Enable=TRUE, premier front toggle IHM -> Diagnostic OK *)
    FB(Enable := TRUE, TglHeartbeatIhm := TRUE, IhmTimeout := T#2s);
    ASSERT_TRUE(FB.HeartbeatIhmOk, 'Enable=TRUE + edge -> HeartbeatIhmOk=TRUE');
    ASSERT_FALSE(FB.HeartbeatIhmTimeout, 'HeartbeatIhmTimeout=FALSE');

    ADVANCE_TIME(10000000);

    (* Scan 2 : Enable=FALSE -> Re-neutralisation *)
    FB(Enable := FALSE, TglHeartbeatIhm := TRUE, IhmTimeout := T#2s);
    ASSERT_FALSE(FB.HeartbeatIhmOk, 'Coupure -> HeartbeatIhmOk retombe a FALSE');
    ASSERT_TRUE(FB.HeartbeatIhmTimeout, 'Coupure -> Timeout=TRUE');
END_TEST

TEST 'TC-P12-020 IHM Heartbeat : surveillance timeout apres 2s sans front'
    (* 1. Initialisation avec front IHM *)
    FB(Enable := TRUE, TglHeartbeatIhm := TRUE, IhmTimeout := T#2s);
    ASSERT_TRUE(FB.HeartbeatIhmOk, 'Heartbeat IHM valide initialement');
    ASSERT_FALSE(FB.HeartbeatIhmTimeout, 'Pas de timeout');

    (* 2. Scan suivant : pas de front, le timer de surveillance démarre *)
    FB(Enable := TRUE, TglHeartbeatIhm := TRUE, IhmTimeout := T#2s);

    (* 3. Avance dans le temps de 2.5s sans nouveau front *)
    ADVANCE_TIME(2500000000);
    FB(Enable := TRUE, TglHeartbeatIhm := TRUE, IhmTimeout := T#2s);
    ASSERT_FALSE(FB.HeartbeatIhmOk, 'Heartbeat IHM tombe en echec apres timeout');
    ASSERT_TRUE(FB.HeartbeatIhmTimeout, 'HeartbeatIhmTimeout leve');

    (* 4. Reprise du toggle IHM -> Retabli *)
    ADVANCE_TIME(10000000);
    FB(Enable := TRUE, TglHeartbeatIhm := FALSE, IhmTimeout := T#2s);
    ASSERT_TRUE(FB.HeartbeatIhmOk, 'Heartbeat IHM retabli apres nouveau front');
    ASSERT_FALSE(FB.HeartbeatIhmTimeout, 'HeartbeatIhmTimeout retombe a FALSE');
END_TEST

(* =========================================================================
   AF-12 — Diagnostic : TC-P12-050 (timeout -> HeartbeatIhmTimeout + TimeSinceIhmEdge)
   ========================================================================= *)

TEST 'TC-P12-050 IHM Heartbeat : timeout -> HeartbeatIhmTimeout + TimeSinceIhmEdge, reprise sur front'
    (* 1. Front IHM initial -> OK *)
    FB(Enable := TRUE, TglHeartbeatIhm := TRUE, IhmTimeout := T#2s, PlcTogglePeriod := T#500ms);
    ASSERT_TRUE(FB.HeartbeatIhmOk, 'Front initial -> HeartbeatIhmOk=TRUE');
    ASSERT_FALSE(FB.HeartbeatIhmTimeout, 'Pas de timeout');

    (* 2. Scan suivant sans front -> timer de surveillance demarre *)
    FB(Enable := TRUE, TglHeartbeatIhm := TRUE, IhmTimeout := T#2s, PlcTogglePeriod := T#500ms);

    (* 3. Avance 2.5s sans front -> timeout, TimeSinceIhmEdge = IhmTimeout *)
    ADVANCE_TIME(2500000000);
    FB(Enable := TRUE, TglHeartbeatIhm := TRUE, IhmTimeout := T#2s, PlcTogglePeriod := T#500ms);
    ASSERT_TRUE(FB.HeartbeatIhmTimeout, 'Timeout apres 2s sans front');
    ASSERT_FALSE(FB.HeartbeatIhmOk, 'HeartbeatIhmOk=FALSE sous timeout');
    ASSERT_EQ(FB.TimeSinceIhmEdge, T#2s, 'TimeSinceIhmEdge = IhmTimeout (2s)');

    (* 4. Nouveau front -> restaure immediatement, TimeSinceIhmEdge repart de 0 *)
    ADVANCE_TIME(10000000);
    FB(Enable := TRUE, TglHeartbeatIhm := FALSE, IhmTimeout := T#2s, PlcTogglePeriod := T#500ms);
    ASSERT_TRUE(FB.HeartbeatIhmOk, 'Nouveau front -> HeartbeatIhmOk restaure');
    ASSERT_FALSE(FB.HeartbeatIhmTimeout, 'Timeout retombe');
    ASSERT_EQ(FB.TimeSinceIhmEdge, T#0s, 'TimeSinceIhmEdge repart de 0');
END_TEST
